    def _pestana_proceso(self):
        pagina = QWidget()
        capa = QHBoxLayout(pagina)
        self.sinoptico = Sinoptico()
        self.sinoptico.accionado.connect(self._accionar)
        capa.addWidget(self.sinoptico, 3)
        caja = QGroupBox("Paradas")
        columna = QVBoxLayout(caja)
        columna.addWidget(rotulo("Clic en pulsadores, cortinas y puerta para simularlos."))
        self.et_paro = QLabel()
        self.et_paro.setWordWrap(True)
        columna.addWidget(self.et_paro)
        self.bt_rearme = QPushButton("Rearme")
        self.bt_rearme.clicked.connect(lambda: self._orden(Op.REARME, self.et_paro_resultado))
        columna.addWidget(self.bt_rearme)
        self.bt_recuperar = QPushButton("Recuperar")
        self.bt_recuperar.clicked.connect(self._recuperar)
        columna.addWidget(self.bt_recuperar)
        self.bt_reiniciar = QPushButton("Reiniciar lote")
        self.bt_reiniciar.clicked.connect(self._reiniciar)
        columna.addWidget(self.bt_reiniciar)
        self.et_paro_resultado = QLabel()
        self.et_paro_resultado.setWordWrap(True)
        columna.addWidget(self.et_paro_resultado)
        columna.addStretch(1)
        capa.addWidget(caja, 1)
        return pagina

    def _pestana_sensores(self):
        pagina = QWidget()
        capa = QVBoxLayout(pagina)
        self.tb_sensores = tabla(("Sensor", "Valor", "Procedencia"))
        capa.addWidget(self.tb_sensores)
        return pagina

    def _pestana_registro(self):
        pagina = QWidget()
        capa = QVBoxLayout(pagina)
        self.tb_registro = tabla(("Fecha", "Usuario", "Perfil", "Operación", "Detalle", "Resultado"))
        capa.addWidget(self.tb_registro)
        return pagina

    def _pestana_administracion(self):
        pagina = QWidget()
        capa = QHBoxLayout(pagina)
        izquierda = QVBoxLayout()
        self.tb_cuentas = tabla(("Usuario", "Nombre", "Perfil", "Activa", "Clave de fábrica"))
        izquierda.addWidget(self.tb_cuentas)
        acciones = QHBoxLayout()
        for texto, funcion in (("Habilitar o inhabilitar", self._alternar_cuenta),
                               ("Cambiar perfil", self._cambiar_perfil),
                               ("Restablecer contraseña", self._restablecer)):
            boton = QPushButton(texto)
            boton.clicked.connect(funcion)
            acciones.addWidget(boton)
        izquierda.addLayout(acciones)
        capa.addLayout(izquierda, 3)
        caja = QGroupBox("Nueva cuenta")
        formulario = QFormLayout(caja)
        self.in_nuevo = QLineEdit()
        self.in_nombre = QLineEdit()
        self.cb_perfil = QComboBox()
        self.cb_perfil.addItems(PERFILES)
        self.in_inicial = QLineEdit()
        self.in_inicial.setEchoMode(QLineEdit.Password)
        formulario.addRow("Usuario", self.in_nuevo)
        formulario.addRow("Nombre", self.in_nombre)
        formulario.addRow("Perfil", self.cb_perfil)
        formulario.addRow("Contraseña", self.in_inicial)
        crear = QPushButton("Crear cuenta")
        crear.setObjectName("crear_cuenta")
        crear.clicked.connect(self._crear_cuenta)
        formulario.addRow(crear)
        self.et_admin = QLabel()
        self.et_admin.setWordWrap(True)
        formulario.addRow(self.et_admin)
        capa.addWidget(caja, 2)
        return pagina

    def _construir_pestanas(self):
        self.pag_proceso = self._pestana_proceso()
        self.pag_produccion = self._pestana_produccion()
        self.pag_mantenimiento = self._pestana_mantenimiento()
        self.pag_sensores = self._pestana_sensores()
        self.pag_registro = self._pestana_registro()
        self.pag_administracion = self._pestana_administracion()

    def _ayuda(self):
        # Solo lista las claves que siguen vigentes: al actualizarlas dejan de mostrarse.
        vigentes = [c["usuario"] for c in self.cuentas.listar()
                    if c["clave_por_defecto"] and c["activo"]]
        cuentas = ("<ul>" + "".join(f"<li><code>{u}</code> / <code>{u}</code></li>" for u in vigentes)
                   + "</ul><p>Actualizarlas al pasar la celda a operación.</p>") if vigentes else \
            "<p>Las contraseñas de fábrica ya fueron actualizadas.</p>"
        self.dialogo_ayuda = QDialog(self)
        self.dialogo_ayuda.setWindowTitle("Ayuda")
        self.dialogo_ayuda.resize(620, 620)
        capa = QVBoxLayout(self.dialogo_ayuda)
        texto = QTextBrowser()
        texto.setHtml(AYUDA.format(cuentas=cuentas))
        capa.addWidget(texto)
        self.dialogo_ayuda.show()

    # Sesión

    def _entrar(self):
        sesion = self.cuentas.autenticar(self.in_usuario.text().strip(), self.in_clave.text())
        self.in_clave.clear()
        if sesion is None:
            self.et_login.setText(FALLO_ACCESO)
            return
        self.sesion = sesion
        self.et_login.clear()
        self.in_usuario.clear()
        self._refrescar_sesion()

    def _cerrar_sesion(self, motivo):
        self.procesador.cerrar_sesion(self.sesion, motivo)
        self.sesion = None
        self.et_login.setText(motivo + ".")
        self._refrescar_sesion()

    def _vigilar_sesion(self):
        if self.sesion is not None and not self.cuentas.sesion_valida(self.sesion):
            self._cerrar_sesion("Sesión cerrada por inactividad o cambio de la cuenta")

    def eventFilter(self, objeto, evento):
        if evento.type() in (QEvent.MouseButtonPress, QEvent.KeyPress):
            self.cuentas.actividad(self.sesion)
        return False

    def _refrescar_sesion(self):
        self.pestanas.clear()
        hay = self.sesion is not None
        self.paginas.setCurrentIndex(1 if hay else 0)
        self.bt_salir.setVisible(hay)
        self.bt_clave.setVisible(hay)
        self.et_usuario.setText(f"{self.sesion.nombre} · {self.sesion.perfil}" if hay else "Sin sesión")
        if hay:
            perfil = self.sesion.perfil
            self.pestanas.addTab(self.pag_proceso, "Proceso")
            self.bt_rearme.setVisible(permitido(perfil, Op.REARME))
            self.bt_recuperar.setVisible(permitido(perfil, Op.RECUPERAR))
            self.bt_reiniciar.setVisible(permitido(perfil, Op.REINICIAR))
            if permitido(perfil, Op.ARRANQUE):
                self.pestanas.addTab(self.pag_produccion, "Producción")
            if permitido(perfil, Op.PREPARAR_MODO):
                self.pestanas.addTab(self.pag_mantenimiento, "Mantenimiento")
            if permitido(perfil, Op.ADMINISTRAR):
                self.pestanas.addTab(self.pag_administracion, "Administración")
            self.pestanas.addTab(self.pag_sensores, "Sensores")
            self.pestanas.addTab(self.pag_registro, "Registro")
            self._refrescar_tablas()
        self._refrescar_aviso()

    def _refrescar_aviso(self):
        texto = ""
        if not self.estado.get("conectado"):
            texto = "Sin conexión con RoboDK: los mandos están bloqueados."
        elif not self.estado.get("estacion_ok"):
            texto = "La estación activa de RoboDK no es la v05: los mandos están bloqueados."
        elif self.estado.get("senales", {}).get("PARO_CAUSA"):
            causa = int(self.estado["senales"]["PARO_CAUSA"])
            texto = f"Celda detenida: {CAUSAS_PARO.get(causa, causa)}. Eliminar la causa y pulsar Rearme."
        elif not self.estado.get("coordinador"):
            texto = "El coordinador está detenido: doble clic en Coordinador_Panel, en RoboDK."
        elif self.estado.get("senales", {}).get("RECUP_PENDIENTE") == 1:
            texto = "Recuperación pendiente: pulsar Recuperar con el perfil de mantenimiento."
        elif self.sesion is not None and self.sesion.clave_por_defecto:
            texto = "Esta cuenta usa la contraseña de fábrica: actualizarla al pasar la celda a operación."
        elif self.sesion is not None and self.sesion.perfil == ADMINISTRADOR \
                and self.cuentas.hay_claves_por_defecto():
            texto = "Hay cuentas con la contraseña de fábrica: actualizarlas al pasar la celda a operación."
        self.aviso.setText(texto)
        self.aviso.setVisible(bool(texto))

    def _refrescar_tablas(self):
        filas = []
        for f in self.cuentas.leer_registro():
            fecha = datetime.fromtimestamp(f["fecha"]).strftime("%d/%m %H:%M:%S")
            filas.append((fecha, f["usuario"], f["perfil"], f["operacion"], f["detalle"], f["resultado"]))
        llenar(self.tb_registro, filas)
        if self.sesion is not None and self.sesion.perfil == ADMINISTRADOR:
            llenar(self.tb_cuentas, [(c["usuario"], c["nombre"], c["perfil"],
                                      "Sí" if c["activo"] else "No",
                                      "Sí" if c["clave_por_defecto"] else "No")
                                     for c in self.cuentas.listar()])

    # Órdenes

    def confirmar(self, texto):
        respuesta = QMessageBox.question(self, "Confirmar", texto, QMessageBox.Yes | QMessageBox.No,
                                         QMessageBox.No)
        return respuesta == QMessageBox.Yes

    def _orden(self, op, etiqueta=None, **datos):
        resultado = self.procesador.solicitar(self.sesion, op, **datos)
        if etiqueta is not None:
            etiqueta.setText(resultado.mensaje)
        elif not resultado.aceptada:
            self.et_login.setText(resultado.mensaje)
        self.cuentas.actividad(self.sesion)
        if self.sesion is not None:
            self._refrescar_tablas()
        return resultado

    def _alternar_emergencia(self):
        pulsada = self.estado.get("senales", {}).get("EMERGENCIA_SIM") == 1
        self._orden(Op.EMERGENCIA, valor=0 if pulsada else 1)

    def _accionar(self, nombre):
        s = self.estado.get("senales", {})
        if nombre == "emergencia":
            self._alternar_emergencia()
            return
        senal = {"cortina_entrada": "CORTINA_ENTRADA_SIM", "cortina_salida": "CORTINA_SALIDA_SIM",
                 "puerta": "PUERTA_ABIERTA_SIM"}[nombre]
        self._orden(Op.RESGUARDO, self.et_paro_resultado, senal=senal, valor=0 if s.get(senal) == 1 else 1)

    def _recuperar(self):
        if self.confirmar("¿Retomar la pieza interrumpida? Los robots van a moverse. Nadie debe estar "
                          "dentro de la zona de robots."):
            self._orden(Op.RECUPERAR, self.et_paro_resultado)

    def _reiniciar(self):
        if self.confirmar("¿Reiniciar el lote? La cinta evacúa, se reponen las piezas y los contadores "
                          "vuelven a cero."):
            self._orden(Op.REINICIAR, self.et_paro_resultado)

    def _preparar(self):
        modo = self.cb_modo.currentData()
        if self.confirmar(f"¿Preparar «{MODOS[modo]}»? Si hay producción, se detendrá al terminar "
                          "la pieza. Nadie debe estar dentro de la zona de robots."):
            self._orden(Op.PREPARAR_MODO, self.et_modo, modo=modo, tipo=self.cb_tipo.currentText())

    def _regresar(self):
        if self.confirmar("¿Confirmás la restitución? Se declara terminada la intervención, con "
                          "resguardos cerrados y nadie dentro. No arranca la producción."):
            self._orden(Op.REGRESAR_MODO, self.et_modo)

    def _entrada(self, senal, marcada):
        self._orden(Op.ENTRADA_SIMULADA, self.et_modo, senal=senal, valor=int(marcada))

    def _cuenta_seleccionada(self):
        fila = self.tb_cuentas.currentRow()
        if fila < 0:
            self.et_admin.setText("Seleccioná una cuenta.")
            return None
        return self.tb_cuentas.item(fila, 0).text()

    def _administrar(self, accion, usuario, *argumentos):
        self.et_admin.setText(self.procesador.administrar(self.sesion, accion, usuario, *argumentos).mensaje)
        self._refrescar_tablas()

    def _crear_cuenta(self):
        self._administrar("crear", self.in_nuevo.text().strip(), self.in_nombre.text().strip(),
                          self.cb_perfil.currentText(), self.in_inicial.text())
        self.in_inicial.clear()

    def _alternar_cuenta(self):
        usuario = self._cuenta_seleccionada()
        if usuario:
            activa = self.tb_cuentas.item(self.tb_cuentas.currentRow(), 3).text() == "Sí"
            self._administrar("habilitar", usuario, not activa)

    def _cambiar_perfil(self):
        usuario = self._cuenta_seleccionada()
        if usuario:
            perfil, ok = QInputDialog.getItem(self, "Cambiar perfil", usuario, PERFILES, 0, False)
            if ok:
                self._administrar("cambiar_perfil", usuario, perfil)

    def _restablecer(self):
        usuario = self._cuenta_seleccionada()
        if usuario:
            clave, ok = QInputDialog.getText(self, "Restablecer contraseña", usuario, QLineEdit.Password)
            if ok:
                self._administrar("fijar_clave", usuario, clave)

    def _cambiar_clave(self):
        actual, ok = QInputDialog.getText(self, "Cambiar contraseña", "Contraseña actual",
                                          QLineEdit.Password)
        if not ok:
            return
        nueva, ok = QInputDialog.getText(self, "Cambiar contraseña", "Contraseña nueva",
                                         QLineEdit.Password)
        if not ok:
            return
        try:
            self.cuentas.cambiar_clave_propia(self.sesion, actual, nueva)
            self.cuentas.registrar(self.sesion.usuario, self.sesion.perfil, "Cambio de contraseña",
                                   "-", "Hecho")
            QMessageBox.information(self, "Contraseña", "Contraseña actualizada.")
        except ErrorCuenta as error:
            QMessageBox.warning(self, "Contraseña", str(error))
        self._refrescar_aviso()

    # Estado

    def recibir_estado(self, estado):
        conectado_antes = self.estado.get("conectado")
        self.estado = estado
        self.procesador.actualizar(estado)
        if conectado_antes and not estado.get("conectado") and self.sesion is not None:
            self._cerrar_sesion("Sesión cerrada por pérdida de conexión")
        s = estado.get("senales", {})
        puerto = estado.get("puerto")
        self.et_conexion.setText(f"RoboDK {puerto}" if estado.get("conectado") else "Sin conexión")
        listo = operativo(estado)
        self.bt_parada.setEnabled(listo)
        self.bt_emergencia.setEnabled(bool(estado.get("conectado") and estado.get("estacion_ok")))
        self.bt_emergencia.setText("LIBERAR EMERGENCIA" if s.get("EMERGENCIA_SIM") == 1 else "EMERGENCIA")
        self.sinoptico.actualizar(s)
        # Stop no pasa por el coordinador: sus señales quedan como estaban y no describen la celda.
        causa_paro = int(s.get("PARO_CAUSA") or 0)
        if causa_paro:
            estado_celda = "Parada: " + CAUSAS_PARO.get(causa_paro, str(causa_paro))
        elif s and not estado.get("coordinador"):
            estado_celda = "Coordinador detenido"
        else:
            estado_celda = ESTADOS.get(int(s.get("ESTADO_CONTROL") or 0), "—") if s else "—"
        self.valores["estado"].setText(estado_celda)
        if not s:
            self.valores["modo"].setText("—")
            self.valores["pieza"].setText("—")
            self.valores["causa"].setText("—")
        else:
            confirmado = int(s.get("MODO_CONFIRMADO") or 0)
            en_transicion = s.get("MODO_EN_TRANSICION") == 1
            self.valores["modo"].setText("Cambiando…" if en_transicion else
                                         MODOS.get(confirmado, "Producción"))
            activa = int(s.get("PIEZA_ACTIVA") or 0)
            proxima = int(s.get("PROXIMA_PIEZA") or 1)
            lote = int(s.get("LOTES_COMPLETADOS") or 0) + 1
            fase = FASES.get(int(s.get("FASE_PIEZA") or 0))
            texto = (f"Lote {lote} · Pieza {activa} de 4" if activa else
                     f"Lote {lote} · Fin de lote" if proxima == 5 else
                     f"Lote {lote} · Próxima {proxima} de 4")
            buenas = int(s.get("PIEZAS_BUENAS") or 0)
            objetivo = int(s.get("OBJETIVO_PIEZAS") or 0)
            retrabajo = int(s.get("PIEZAS_RETRABAJO") or 0)
            meta = f"{buenas} de {objetivo} buenas" if objetivo else f"{buenas} buenas"
            detalle = f"{meta} · {retrabajo} retrabajo" + (f" · {fase}" if activa and fase else "")
            self.valores["pieza"].setText(texto + "\n" + detalle)
            causa = int(s.get("CAUSA_RECHAZO") or 0) or int(s.get("MODO_CAUSA") or 0)
            self.valores["causa"].setText(self.causas.get(causa, str(causa)) if causa else "Ninguno")
        self._actualizar_mandos(s, listo)
        self._refrescar_aviso()

    def _actualizar_mandos(self, s, listo):
        if self.sesion is None:
            return
        causa_paro = int(s.get("PARO_CAUSA") or 0)
        self.et_paro.setText(f"Parada activa: {CAUSAS_PARO.get(causa_paro, causa_paro)}" if causa_paro else
                             "Recuperación pendiente" if s.get("RECUP_PENDIENTE") == 1 else "Sin paradas")
        self.bt_rearme.setEnabled(bool(causa_paro))
        self.bt_recuperar.setEnabled(bool(listo and not causa_paro and s.get("RECUP_PENDIENTE") == 1))
        self.bt_reiniciar.setEnabled(bool(listo and not causa_paro and s.get("AUTO_ACTIVO") == 0
                                          and s.get("RECUP_PENDIENTE") == 0))
        condiciones = condiciones_arranque(s)
        faltan = [nombre for nombre, ok in condiciones if not ok]
        automatico = s.get("AUTO_ACTIVO") == 1
        self.et_condiciones.setText("\n".join(f"{'Cumple' if ok else 'Falta '}  ·  {nombre}"
                                              for nombre, ok in condiciones))
        self.bt_arranque.setEnabled(listo and not automatico and not faltan)
        if automatico:
            self.et_arranque.setText("Producción en curso.")
        elif not listo:
            self.et_arranque.setText("Sin conexión con el coordinador.")
        elif faltan:
            self.et_arranque.setText("Falta: " + ", ".join(faltan).lower() + ".")
        else:
            self.et_arranque.setText("Listo para arrancar.")
        confirmado = int(s.get("MODO_CONFIRMADO") or 0)
        libre = listo and s.get("MODO_EN_TRANSICION") == 0
        self.bt_preparar.setEnabled(bool(libre and confirmado == 0))
        self.bt_regresar.setEnabled(bool(libre and confirmado != 0))
        resultado = int(s.get("MODO_RESULTADO") or 0)
        if resultado:
            causa = int(s.get("MODO_CAUSA") or 0)
            texto = RESULTADOS_MODO.get(resultado, "—")
            self.et_modo.setText(f"Última solicitud: {texto}" +
                                 (f" · {self.causas.get(causa, causa)}" if causa else ""))
        for senal, casilla in self.entradas.items():
            casilla.setEnabled(bool(self.estado.get("conectado") and self.estado.get("estacion_ok")))
            casilla.setChecked(s.get(senal) == 1)
        llenar(self.tb_sensores, [(nombre, "Sí" if s.get(senal) == 1 else "No",
                                   "Calculado por Python") for senal, nombre in SENSORES] +
               [(ETIQUETAS_ENTRADA[e], "Sí" if s.get(e) == 1 else "No", "Entrada simulada")
                for e in ENTRADAS_SIMULADAS])

    def closeEvent(self, evento):
        self.procesador.cerrar_sesion(self.sesion, "Cierre del panel")
        evento.accept()

# --- panel.py ---

def crear(ruta=None, puertos=PUERTOS):
    enlace = Enlace(puertos)
    cuentas = Cuentas(ruta or ruta_datos())
    procesador = Procesador(cuentas, enlace.enviar, CAUSAS)
    ventana = Ventana(cuentas, procesador, CAUSAS)
    enlace.estado.connect(ventana.recibir_estado)
    return enlace, cuentas, procesador, ventana

def main():
    parser = argparse.ArgumentParser()
    parser.add_argument("--puerto", type=int)
    args = parser.parse_args()
    app = QApplication(sys.argv)
    enlace, _, _, ventana = crear(puertos=(args.puerto,) if args.puerto else PUERTOS)
    app.installEventFilter(ventana)
    ventana.show()
    enlace.start()
    codigo = app.exec_()
    enlace.detener()
    sys.exit(codigo)

if __name__ == "__main__":
    main()
